(* IEC 61131-3 sources: rk/crates/fuzz/regressions, 25 files *)

(* ---- format-unparsable--a-case-label-read-as-an-assignment-missing-its-equal.st ---- *)
TYPE STATE: INT(A, B, C) END_TYPE
FUNCTION test : INT
VAR x : STATE; END_VAR
    CASE x OF
        STATE#A: test z:= 10;
        STATE#B: test :CONTINUE+EMENTSTATE#A: test := 02;
ABSTRACT    END_CASE;
END_FUNCTION

(* ---- format-unparsable--pragma-text-dropped.st ---- *)
        TYPE
            Matrix: ARRAY[1..2, 1..3] OF INT{export};
        END_TYPE

        FUNCTION Test
            VAR
                Data : Matrix := [[1, 2, 3], [4, 5, 6], [7, 8, 9]];
            END_VAR
        END_FUNCTION

(* ---- ide-tokens--a-path-before-a-stray-operator.st ---- *)
TYPE
    Step : (A := 5, B, C);
    Holder : STRUCT s : Step; END_STRUCT;
END_TYPE
FUNCTION test : INT
VAR
    h : Holder;
END_VAR
    IF h.s ! Step#A THEN test := test + 1; END_IF;
END_FUNCTION

(* ---- panic--a-repetition-given-as-an-array-field-s-value.st ---- *)
(* `arr` is given a repetition of brackets with no brackets of its own. The
   checks passed it and nothing placed its values, so `m.arr` stayed 0, and
   the assertion that an initializer drops no value panicked. It is E0515. *)

TYPE M : STRUCT arr : ARRAY[0..3] OF INT; END_STRUCT; END_TYPE

FUNCTION F
VAR
    m : M := (arr := 2([1, 2]));
END_VAR
END_FUNCTION

(* ---- edit-text--pasted-junk-cutting-a-crlf-in-two.st ---- *)
        FUNCTION run : DINT
        VAR inner : STRING; outer : STRING; END_VAR
            __TRY
                __TRY
                    __RAISE('first');
                __CATCH(inner)
                    run := 1;
                __END_TRY;
                __TRY
                    __RAISE('second');
                __CATCH(inner)
                    __RAISE(inner);
                __END_TRY;
  + 10;
                END_IF;
            __END_TRY;
        END_FUN/*ION

(* ---- format-idempotence--an-extern-pragma-over-two-lines.st ---- *)
FUNCTION B : INT
END_FUNCTION{
extern 'm' 'n'}
FUNCTION C : INT
END_FUNCTION

(* ---- ide-edits--a-namespace-named-for-several-variables.st ---- *)
    FUNCTION fn1
    VAR
        counter, y : INPROT.CTEDD_VAR
        counter += 2;
        y := counter := 1;
        counter *= coRESOURCEunter;
        y += counter -= 1;
        counter += y := counter;
    END_FUNCTION

(* ---- ide-range--a-related-label-in-the-library.st ---- *)
FUNCTION f : DINT
VAR CONSTANT
    N : DINT := 200 * 200;
    HALF : INT := 20000;
END_VAR
VAR
    x : DINT;
END_VAR
    x := 32767 + 1;
    x := INT#200 * INT#200;
    x := (HALF * 2) + 1;
    f := N;
END_FUNCTION

(* ---- incremental-parse--comments-shifted-after-closing-one.st ---- *)
FUNCTION f : INT
VAR
    x : INT; // one
    y : INT; (* two *)
END_VAR // after the section
    x := 1; // one
    y := 2; (* two *)
    IF x = 1 THEN // why
        x := 3; // three
        // alone
    ELSE // other
        x := 4;
    END_IF; // closed
    // alone again
    f := x; /* last */
END_FUNCTION // done

(* ---- panic--an-initializer-of-an-unknown-type.st ---- *)
(* `Point` and `Holder` are declared nowhere. Past an unknown type the walk
   says nothing more and places nothing, and the assertion that no value is
   dropped panicked on a program that never compiles. *)

FUNCTION f
VAR
    rows : ARRAY[0..1] OF Point := [(1, 2), (3, 4)];
    nested : Holder := (p := (y := 3, 4), 5);
END_VAR
END_FUNCTION

(* ---- profiles-diverge--a-test-function.st ---- *)
{test}
FUNCTION my_test : INT
END_FUNCTION

(* ---- format-meaning--the-formatted-text-read-with-other-addresses.st ---- *)
        TYPE Tally : INT := 5; END_TYPE
        TYPE B8 : BYTE := 16#FF; END_TYPE

        FUNCTION_BLOCK Drive
        VAR
            m AT %M* : Tally;
            b AT %Q* : B8;
            c AT %M* : Tally;
        END_VAR
        END_FUNCTION_BLOCK

        PROGRAM P
        VAR d : Drive; END_VAR
            d();
        END_PROGRAM

        CONFIGURATION Cfg
        VAR_GLOBAL
            g AT %MW0 : INT := 7;
            w AT %QD0 : DWORD := 16#11223344;
        END_VAR
        VAR_CONFIG
            Res.P1.d.m AT %MW0 : Tally;
            Res.P1.d.b AT %QB2 : B8;
            Res.P1.d.c AT %MW1 : Tally;
        END_VAR
            RESOURCE Res ON CPU
                TASK T(INTERVAL := T#10ms, PRIORITY := 1);
                PROGRAM P1 WITH T : P;
            END_RESOURCE
        END_CONFIGURATION

// v2

(* ---- ide-range--a-definition-in-the-library.st ---- *)
        TYPE Holder : STRUCT p : REF_TO INT; END_STRUCT; END_TYPE

        FUNCTION test : INT
        VAR
            x : INT :=D_TYPE

        FUNCTION_BLOCK Holder
        VAR_OUTPUT r : REAL; END_VAR
        END_FUNCTION_BLOCK

        FUNCTION Half : REAL
            Half := 0.5;
            Half.31 := TRUE; 42;
            h : Holder := (p := REF(x));
        END_VAR
            test := h.p^;
        END_NCTCTION

(* ---- lowering--a-real-constant-computed-from-another-as-an-initial-value.st ---- *)
(* rk-fuzz expects, after 1 scans:
P1.f.m = 3.0
g = 3.0
*)

FUNCTION_BLOCK Fb
VAR CONSTANT
    k0 : REAL := 1.5;
    k1 : REAL := k0 * 2.0;
END_VAR
VAR
    m : REAL := k1;
END_VAR
END_FUNCTION_BLOCK

PROGRAM Main
VAR
    f : Fb;
END_VAR
    f();
END_PROGRAM

CONFIGURATION Cfg
    VAR_GLOBAL CONSTANT
        g0 : REAL := 1.5;
        g1 : REAL := g0 * 2.0;
    END_VAR
    VAR_GLOBAL
        g : REAL := g1;
    END_VAR
    RESOURCE R ON CPU
        TASK T(INTERVAL := T#10ms, PRIORITY := 1);
        PROGRAM P1 WITH T : Main;
    END_RESOURCE
END_CONFIGURATION

(* ---- panic--a-member-value-repeated-without-its-parentheses.st ---- *)
(* The standard's table of user-defined types gives each instance of an array
   of TON its PT with a repetition of the member value, which has no
   parentheses of its own. The checks passed it, nothing placed PT, and the
   assertion that no value is dropped panicked. Each instance gets it now. *)

FUNCTION_BLOCK Timer
VAR_INPUT PT : TIME; END_VAR
END_FUNCTION_BLOCK

TYPE Timers : ARRAY[1..20] OF Timer := [20(PT := T#250ms)]; END_TYPE

PROGRAM P
VAR t : Timers; END_VAR
    t[1]();
END_PROGRAM

(* ---- panic--implements-before-an-extends-with-no-base.st ---- *)
INTERFACE ITF1
    METHOD DoWork END_METHOD
END_INTERFACE

FUNCTION_BLOCK Impl IMPLEMENTS ITF1
   EXTENDS METHOD DoWork END_METHOD
END_FUNCTION_BLOCK

FUNCTION Use : INT
    VAR_IN_OUT dev : ITF1; END_VAR
    VAR other : Impl; END_VAR
    dev := other;
END_FUNCTION

(* ---- semantics--a-member-named-like-another-type.st ---- *)
(* rk-fuzz expects, after 1 scans:
P1.f.out = 2
P1.f.e1 = 5
*)

TYPE E0 : INT (n0 := 5, n1 := 7);
END_TYPE

TYPE E1 : INT (n0 := 1, n1 := 2);
END_TYPE

FUNCTION_BLOCK fb
VAR
    e1 : E0 := E0#n0;
END_VAR
VAR_OUTPUT
    out : INT;
END_VAR
    out := E1#n1;
END_FUNCTION_BLOCK

PROGRAM Main
VAR
    f : fb;
END_VAR
    f();
END_PROGRAM

CONFIGURATION Cfg
    RESOURCE R ON CPU
        TASK T(INTERVAL := T#10ms, PRIORITY := 1);
        PROGRAM P1 WITH T : Main;
    END_RESOURCE
END_CONFIGURATION

(* ---- spacing--the-base-body-s-call-with-spaced-parentheses.st ---- *)
FUNCTION_BLOCK base
END_FUNCTION_BLOCK

FUNCTION_BLOCK spaced_inside EXTENDS base
    SUPER(		);
END_FUNCTION_BLOCK

FUNCTION_BLOCK spaced_before EXTENDS base
    SUPER ( );
END_FUNCTION_BLOCK

(* ---- ide-edits--a-namespace-around-a-recovered-name.st ---- *)
NAMESPACE b
    NAMESPACE a ...args
    END_NAMESPACE
END_NAMESPACE

(* ---- incremental-parse--comment-shifted-after-a-deletion.st ---- *)
        PROGRAM P
        VAR RETAIN seen : STRING[10]; END_VAR
        VAR src : STRING[8]; END_VAR
            src := 'abcdef';
            g := src;   (* from a variable: an over-long literal is E0306 *)
            seen := g;
        END_PROGRAM

        CONFIGURATION Cfg
        VAR_GLOBAL g : STRING[4]; END_VAR
            RESOURCE Res ON CPU
                TASK T(INTERVAL := T#10ms, PRIORITY := 1);
                PROGRAM P1 WITH T : P;
            END_RESOURCE
        END_CONFIGURATION

(* ---- lowering--a-case-label-that-is-a-constant-of-a-named-values-type.st ---- *)
(* rk-fuzz expects, after 1 scans:
P1.hit = 1
*)

TYPE Light : INT (Red := 1, Amber := 2, Green := 3);
END_TYPE

PROGRAM Main
VAR CONSTANT
    k : Light := Light#Amber;
END_VAR
VAR
    m : Light := Light#Amber;
    hit : INT;
END_VAR
    CASE m OF
        k: hit := 1;
    ELSE
        hit := 2;
    END_CASE;
END_PROGRAM

CONFIGURATION Cfg
    RESOURCE R ON CPU
        TASK T(INTERVAL := T#10ms, PRIORITY := 1);
        PROGRAM P1 WITH T : Main;
    END_RESOURCE
END_CONFIGURATION

(* ---- lowering--a-power-in-a-value-init-stores.st ---- *)
(* rk-fuzz expects, after 1 scans:
P1.p = 2.25
g = 8.0
*)

PROGRAM Main
VAR
    p : REAL := 1.5 ** 2.0;
END_VAR
    p := p;
END_PROGRAM

CONFIGURATION Cfg
    VAR_GLOBAL CONSTANT
        k : REAL := 3.0;
    END_VAR
    VAR_GLOBAL
        g : REAL := 2.0 ** k;
    END_VAR
    RESOURCE R ON CPU
        TASK T(INTERVAL := T#10ms, PRIORITY := 1);
        PROGRAM P1 WITH T : Main;
    END_RESOURCE
END_CONFIGURATION

(* ---- lowering--a-reference-compared-with-a-ref.st ---- *)
TYPE
    Row : ARRAY[0..1] OF INT;
END_TYPE

PROGRAM Main
VAR
    l : LINT;
    x : REAL;
    s : STRING;
    row : Row;
    rl : REF_TO LINT;
    rx : REF_TO REAL;
    rs : REF_TO STRING;
    rrow : REF_TO Row;
    a, b, c, d : BOOL;
END_VAR
    rl := REF(l);
    rx := REF(x);
    rs := REF(s);
    rrow := REF(row);
    a := rl = REF(l);
    b := REF(x) = rx;
    c := rs <> REF(s);
    d := rrow = REF(row);
END_PROGRAM

CONFIGURATION Cfg
    RESOURCE Res ON CPU
        TASK T(INTERVAL := T#10ms, PRIORITY := 1);
        PROGRAM P1 WITH T : Main;
    END_RESOURCE
END_CONFIGURATION

(* ---- lowering--a-slice-through-a-path-bound-to-an-in-out.st ---- *)
TYPE
    Rec : STRUCT w : WORD; END_STRUCT;
END_TYPE

FUNCTION set_it
VAR_IN_OUT v : BOOL; END_VAR
    v := TRUE;
END_FUNCTION

PROGRAM Main
VAR
    rec : Rec;
    list : ARRAY[0..1] OF WORD;
END_VAR
    set_it(rec.w.2);
    set_it(list[1].2);
END_PROGRAM

CONFIGURATION Cfg
    RESOURCE Res ON CPU
        TASK T(INTERVAL := T#10ms, PRIORITY := 1);
        PROGRAM P1 WITH T : Main;
    END_RESOURCE
END_CONFIGURATION

(* ---- panic--a-reference-type-that-comes-back-to-itself.st ---- *)
TYPE
    A : ARRAY[0..1] OF REF_TO A;
    P : REF_TO P;
    Q : REF_TO R;
    R : REF_TO Q;
END_TYPE

PROGRAM Main
VAR
    a1, a2 : A;
    p1, p2 : P;
    q1 : Q;
    r1 : R;
    same : BOOL;
END_VAR
    a1[0] := REF(a2);
    a1[0]^[1] := REF(a1);
    p1 := REF(p2);
    p2 := p1;
    q1 := REF(r1);
    r1 := REF(q1);
    same := q1^ = r1;
END_PROGRAM

CONFIGURATION Cfg
    RESOURCE Res ON CPU
        TASK T(INTERVAL := T#10ms, PRIORITY := 1);
        PROGRAM P1 WITH T : Main;
    END_RESOURCE
END_CONFIGURATION
